(* PLC project , CODESYS CODESYS V3.5 SP16 Patch 4 *)
(* stored: creationDateTime 2021-05-05T17:51:35.7556752, modificationDateTime 2021-05-05T17:51:02.9781549 *)

FUNCTION_BLOCK hvac_logic
  VAR_INPUT
    HVAC_ACK : BOOL;
    HVAC_RQ : BOOL;
    HVAC_IN : BOOL;
    HVAC_BYPASS : BOOL;
  END_VAR
  VAR_OUTPUT
    HVAC_RN : BOOL;
    HVAC_STATUS_EN : BOOL;
    HVAC_STATUS_RQ : BOOL;
  END_VAR
  VAR
    TON_0 : TON;
    TON_1 : TON;
    TON_1_ET : TIME;
  END_VAR
  VAR CONSTANT
    HVAC_TIME : TIME := TIME#14ms;
  END_VAR

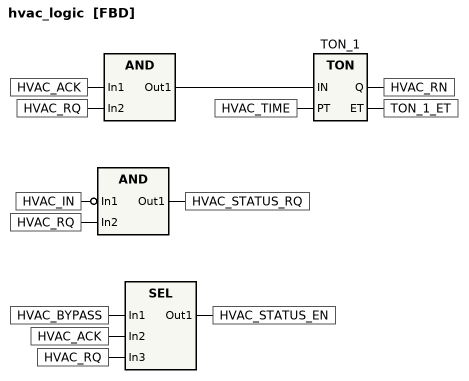
(* FBD diagram, written out as Structured Text *)
TON_1(IN := HVAC_ACK AND HVAC_RQ, PT := HVAC_TIME, ET => TON_1_ET);
HVAC_RN := TON_1.Q;
HVAC_STATUS_RQ := NOT HVAC_IN AND HVAC_RQ;
HVAC_STATUS_EN := SEL(HVAC_BYPASS, HVAC_ACK, HVAC_RQ);
END_FUNCTION_BLOCK
